Fanuc KAREL source: KB00155.KL

PROGRAM KB00155
%NOLOCKGROUP
%ENVIRONMENT MEMO
VAR
  P1: STRING[80]
  P2: INTEGER
BEGIN
  P1 = 'A'
  P2 = 1
  SAVE_DRAM(P1, P2)
END KB00155
